(* IEC 61131-3 sources: PLC-Static-Analysis/modules/plc-rules/src/test/resources/PLCA-Q008/tasks, 1 file *)

(* ---- project.st ---- *)
PROGRAM P_Fast
END_PROGRAM

PROGRAM P_Test // PLCA-Q008
END_PROGRAM

CONFIGURATION Cfg
    RESOURCE Res ON PLC
        TASK tFast(INTERVAL := T#2MS, PRIORITY := 1);
        PROGRAM iFast WITH tFast : P_Fast;
    END_RESOURCE
END_CONFIGURATION
